FUNCTION_BLOCK T_E_text_Safety EXTENDS T_E_text_Common
VAR
END_VAR

PROPERTY errorDoor_0 : ST_E_Text
GET
errorDoor_0.Number:= 13;
END_GET
END_PROPERTY

PROPERTY errorEStop_0 : ST_E_Text
GET
errorEStop_0.Number:= 12;
END_GET
END_PROPERTY

PROPERTY errorGroupCom : KOSTAL_AF2024_Core_Text.ST_E_Text
GET
errorGroupCom.Number:= 10;
END_GET
END_PROPERTY

PROPERTY errorGroupFb : ST_E_Text
GET
errorGroupFb.Number:= 11;
END_GET
END_PROPERTY

PROPERTY safetyNok : ST_E_Text
GET
safetyNok.Number:= 5;
END_GET
END_PROPERTY

PROPERTY safetyOk : ST_E_Text
GET
safetyOk.Number:= 4;
END_GET
END_PROPERTY

PROPERTY safetyRelay_0 : ST_E_Text
GET
safetyRelay_0.Number:= 14;
END_GET
END_PROPERTY

END_FUNCTION_BLOCK

(* stored: Version 1.1.0.1, ProductVersion 3.1.4024.12
   POU T_E_text_Safety: Id {7ecd4c03-6104-4c78-831d-d794bc761f51}, SpecialFunc None
   Property errorDoor_0: Id {2ef9f95c-e717-4c5a-9f02-2332fee5bbe7}
   Get Get: Id {d2acc0ee-f067-474a-9a5f-139919dfcf29}
   Property errorEStop_0: Id {22ec61af-cc72-4c7d-9085-190c54540a24}
   Get Get: Id {3b60cb18-b979-4679-9db6-8ad6a2d62b3b}
   Property errorGroupCom: Id {51e56854-8778-4d12-8492-5021af1fbff9}
   Get Get: Id {68426aa1-6872-4f7f-bd7e-f5e55f0f2f83}
   Property errorGroupFb: Id {2f1bebaf-00b7-41a9-8e90-dcc77da18832}
   Get Get: Id {099e1515-b1ae-46ac-9cc7-3e206a9cca37}
   Property safetyNok: Id {2e565c95-cc4c-4c5b-97f1-036c5db99d7c}
   Get Get: Id {99bac8a4-ddf6-478d-9765-16dc4e5e91da}
   Property safetyOk: Id {f839acea-d733-465e-be40-bfa31e060e34}
   Get Get: Id {469a4a5c-b19a-49a8-94cd-f217abb251ba}
   Property safetyRelay_0: Id {61dd033c-3085-4e49-896b-39bff657ced4}
   Get Get: Id {583ed0e1-bd49-4246-b329-2e164038cb04} *)
